FUNCTION_BLOCK Testing (* CAT Function Block Type *)
  (* Standard: 61499-2 *)
  (* Version 0.0, 11/16/2026, Sandeep Patil, Flexbridge AB, template *)
  PACKAGE Flexbridge.FestoMPS400;
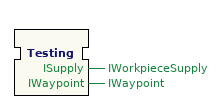
  PLUGS
    ISupply : IWorkpieceSupply;
    IWaypoint : IWaypoint;
  END_PLUGS
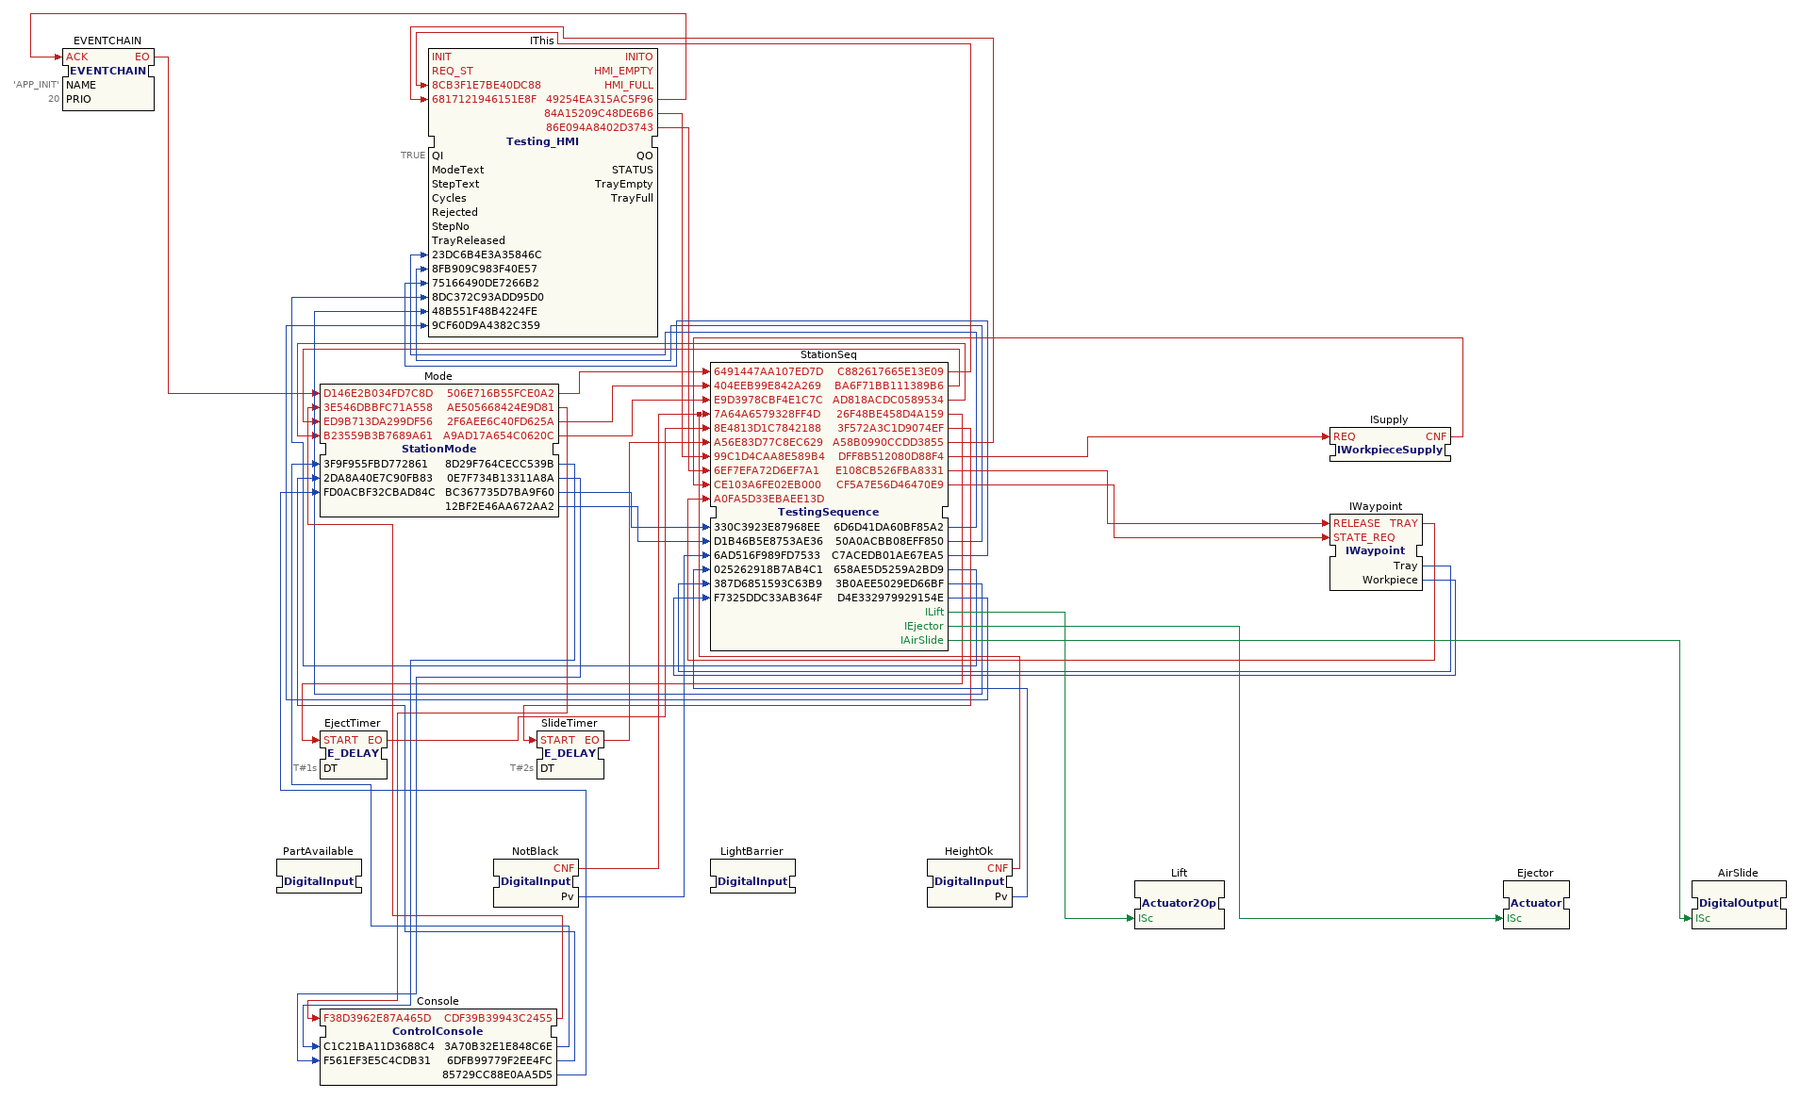
  (* 0 - INITIALIZATION *)
  (* 6 - HMI INTERFACE *)
  (* 1 - FUNCTIONAL INPUT INTERFACE *)
  (* 5 - LOGICS *)
  (* 2 - FUNCTIONAL OUTPUT INTERFACE (ISupply to Distributing, IWaypoint to the conveyor) *)
  (* 3 - FIELD INTERFACE (3.B FROM THE FIELD: sensors, console) *)
  (* 4 - CHILDREN *)
  (* 4.A - TYPICALS (one device CAT per Festo device) *)
  FBS
    Lift : Actuator2Op;
    Ejector : Actuator;
    AirSlide : DigitalOutput;
    PartAvailable : DigitalInput;
    NotBlack : DigitalInput;
    LightBarrier : DigitalInput;
    HeightOk : DigitalInput;
    Console : ControlConsole;
    EVENTCHAIN : EVENTCHAIN(NAME := 'APP_INIT', PRIO := 20);
    IThis : Testing_HMI(QI := TRUE);
    Mode : StationMode;
    StationSeq : TestingSequence;
    EjectTimer : E_DELAY(DT := T#1s);
    SlideTimer : E_DELAY(DT := T#2s);
  END_FBS
  EVENT_CONNECTIONS
    EVENTCHAIN.EO TO Mode.D146E2B034FD7C8D;
    Mode.506E716B55FCE0A2 TO StationSeq.6491447AA107ED7D;
    StationSeq.C882617665E13E09 TO IThis.8CB3F1E7BE40DC88;
    IThis.49254EA315AC5F96 TO EVENTCHAIN.ACK;
    Console.CDF39B39943C2455 TO Mode.3E546DBBFC71A558;
    Mode.AE505668424E9D81 TO Console.F38D3962E87A465D;
    Mode.2F6AEE6C40FD625A TO StationSeq.404EEB99E842A269;
    StationSeq.BA6F71BB111389B6 TO Mode.ED9B713DA299DF56;
    StationSeq.AD818ACDC0589534 TO Mode.B23559B3B7689A61;
    Mode.A9AD17A654C0620C TO StationSeq.E9D3978CBF4E1C7C;
    NotBlack.CNF TO StationSeq.7A64A6579328FF4D;
    HeightOk.CNF TO StationSeq.7A64A6579328FF4D;
    StationSeq.26F48BE458D4A159 TO EjectTimer.START;
    EjectTimer.EO TO StationSeq.8E4813D1C7842188;
    StationSeq.3F572A3C1D9074EF TO SlideTimer.START;
    SlideTimer.EO TO StationSeq.A56E83D77C8EC629;
    StationSeq.A58B0990CCDD3855 TO IThis.6817121946151E8F;
    IThis.84A15209C48DE6B6 TO StationSeq.99C1D4CAA8E589B4;
    IThis.86E094A8402D3743 TO StationSeq.6EF7EFA72D6EF7A1;
    StationSeq.DFF8B512080D88F4 TO ISupply.REQ;
    ISupply.CNF TO StationSeq.CE103A6FE02EB000;
    IWaypoint.TRAY TO StationSeq.A0FA5D33EBAEE13D;
    StationSeq.E108CB526FBA8331 TO IWaypoint.RELEASE;
    StationSeq.CF5A7E56D46470E9 TO IWaypoint.STATE_REQ;
  END_CONNECTIONS
  DATA_CONNECTIONS
    Console.3A70B32E1E848C6E TO Mode.3F9F955FBD772861;
    Console.6DFB99779F2EE4FC TO Mode.2DA8A40E7C90FB83;
    Console.85729CC88E0AA5D5 TO Mode.FD0ACBF32CBAD84C;
    Mode.8D29F764CECC539B TO Console.C1C21BA11D3688C4;
    Mode.0E7F734B13311A8A TO Console.F561EF3E5C4CDB31;
    Mode.BC367735D7BA9F60 TO StationSeq.330C3923E87968EE;
    Mode.12BF2E46AA672AA2 TO StationSeq.D1B46B5E8753AE36;
    NotBlack.Pv TO StationSeq.6AD516F989FD7533;
    HeightOk.Pv TO StationSeq.025262918B7AB4C1;
    IWaypoint.Tray TO StationSeq.387D6851593C63B9;
    IWaypoint.Workpiece TO StationSeq.F7325DDC33AB364F;
    StationSeq.6D6D41DA60BF85A2 TO IThis.23DC6B4E3A35846C;
    StationSeq.50A0ACBB08EFF850 TO IThis.8FB909C983F40E57;
    StationSeq.C7ACEDB01AE67EA5 TO IThis.75166490DE7266B2;
    StationSeq.658AE5D5259A2BD9 TO IThis.8DC372C93ADD95D0;
    StationSeq.3B0AEE5029ED66BF TO IThis.48B551F48B4224FE;
    StationSeq.D4E332979929154E TO IThis.9CF60D9A4382C359;
  END_CONNECTIONS
  ADAPTER_CONNECTIONS
    StationSeq.ILift TO Lift.ISc;
    StationSeq.IEjector TO Ejector.ISc;
    StationSeq.IAirSlide TO AirSlide.ISc;
  END_CONNECTIONS
END_FUNCTION_BLOCK
